(* IEC 61131-3 sources: kns-port-domestic/targets/astra/lib/src/POUs/Util/F_RateLimit, 2 files *)

(* ---- F_RateLimit.decl.st ---- *)
// Назначение: шаг ограничителя скорости изменения: значение движется от rCurrent к rTarget
//             не быстрее rRateUp_ups (рост) и rRateDown_ups (спад) инж. ед. в секунду за шаг
//             lrDt_s. Скорость 0 (или меньше) — без ограничения. lrDt_s <= 0 или rTarget не
//             конечно (NaN из Modbus/ПИД) — значение не меняется. Расчёт шага — в LREAL.
// Автор:      kr0nsch
// Версия:     0.1.0
// Документ:   docs/fb/Functions.md
FUNCTION F_RateLimit : REAL
VAR_INPUT
    rCurrent      : REAL;    // текущее значение (результат прошлого шага)
    rTarget       : REAL;    // цель
    rRateUp_ups   : REAL;    // предел скорости роста, инж. ед./с; <= 0 — без ограничения
    rRateDown_ups : REAL;    // предел скорости спада, инж. ед./с; <= 0 — без ограничения
    lrDt_s        : LREAL;   // шаг времени, с
END_VAR
VAR
    lrLimit : LREAL;         // достижимое за шаг значение
END_VAR

(* ---- F_RateLimit.impl.st ---- *)
IF lrDt_s <= 0.0 OR NOT F_IsFinite(rIn := rTarget) THEN
    // шага нет или цель — мусор: значение не меняется
    F_RateLimit := rCurrent;
ELSIF rTarget > rCurrent AND rRateUp_ups > 0.0 THEN
    // рост, ограничен сверху
    lrLimit := REAL_TO_LREAL(rCurrent) + REAL_TO_LREAL(rRateUp_ups) * lrDt_s;
    F_RateLimit := LREAL_TO_REAL(MIN(REAL_TO_LREAL(rTarget), lrLimit));
ELSIF rTarget < rCurrent AND rRateDown_ups > 0.0 THEN
    // спад, ограничен снизу
    lrLimit := REAL_TO_LREAL(rCurrent) - REAL_TO_LREAL(rRateDown_ups) * lrDt_s;
    F_RateLimit := LREAL_TO_REAL(MAX(REAL_TO_LREAL(rTarget), lrLimit));
ELSE
    // цель достигнута, скорость не ограничена или текущее значение не число: сразу к цели
    F_RateLimit := rTarget;
END_IF
